PROGRAM Test
VAR
	fbEventBufferTest: FB_EventBuffer_Test();
END_VAR

TcUnit.RUN();

END_PROGRAM

(* stored: Version 1.1.0.1
   POU Test: Id {3b6656aa-89b0-446f-8928-0341e81ec3ab}, SpecialFunc None *)
